Omron Sysmac Studio project SF_PLC ver.2 (Sysmac Studio 1.53.0.9, StandardProject)

# Controller new_controller_0: NX102-1020 version 1.33
Units and slaves: 노드1 : NX-ECC203 (E001); 유니트 1 : NX-ID6142-6 (N1); 유니트 2 : NX-OD6121-6 (N2); 유니트 1 : NX-PF0730 (N3); 유니트 2 : NX-ILM400 (N4); 유니트 4 : NX-SID800 (N6); 유니트 5 : NX-SOD400 (N7)
Task PrimaryTask (priority 4, period or condition 2000): Program0

TYPE Robot_IO : STRUCT
    IO : IO16;
END_STRUCT END_TYPE
TYPE IO16 : UNION
    w : WORD;
    b : ARRAY[1..32] OF BOOL;
END_UNION END_TYPE

VAR_GLOBAL
    Robot_In : ARRAY[0..237] OF WORD;  (* 로봇 > PLC; network input *)
    Robot_Out : ARRAY[0..105] OF WORD;  (* PLC > 로봇; network output *)
    vision_trig : BOOL;  (* 비전 촬영 신호; at ECAT://node#4/Line0 Trigger *)
    vis_data : DINT;  (* 비전 데이터; at ECAT://node#4/Line0 DINT Result Data 0 *)
    r_pause : BOOL;  (* 태스크 일시정지; at ECAT://node#[1,2]/Output Bit 32 bits/Output Bit 04 *)
    syl_f : BOOL;  (* 배출 실린더 전진; at ECAT://node#[1,2]/Output Bit 32 bits/Output Bit 05 *)
    syl_r : BOOL;  (* 배출 실린더 후진; at ECAT://node#[1,2]/Output Bit 32 bits/Output Bit 06 *)
    r_resume : BOOL;  (* 태스크 재개; at ECAT://node#[1,2]/Output Bit 32 bits/Output Bit 13 *)
    tower_R : BOOL;  (* 타워램프 - red; at ECAT://node#[1,2]/Output Bit 32 bits/Output Bit 20 *)
    tower_Y : BOOL;  (* 타워램프 - yellow; at ECAT://node#[1,2]/Output Bit 32 bits/Output Bit 21 *)
    tower_G : BOOL;  (* 타워램프 - green; at ECAT://node#[1,2]/Output Bit 32 bits/Output Bit 22 *)
    r_start : BOOL;  (* 태스크 실행; at ECAT://node#[1,2]/Output Bit 32 bits/Output Bit 23 *)
    r_stop : BOOL;  (* 태스크 정지; at ECAT://node#[1,2]/Output Bit 32 bits/Output Bit 24 *)
    vision_ss : BOOL;  (* 비전 감지 센서; at ECAT://node#[1,1]/Input Bit 32 bits/Input Bit 19 *)
    mag_ss : BOOL;  (* 매거진 센서; at ECAT://node#[1,1]/Input Bit 32 bits/Input Bit 23 *)
    stop_ss : BOOL;  (* 스토퍼 센서; at ECAT://node#[1,1]/Input Bit 32 bits/Input Bit 24 *)
    rsol_ss : BOOL;  (* 실린더 후진 센서; at ECAT://node#[1,1]/Input Bit 32 bits/Input Bit 25 *)
    fsol_ss : BOOL;  (* 실린더 전진 센서; at ECAT://node#[1,1]/Input Bit 32 bits/Input Bit 26 *)
    m_run : WORD;  (* 모터 구동; at ECAT://node#2/Command *)
    m_vel : UINT := 5000;  (* 모터 속도; at ECAT://node#2/Frequency reference *)
    m_status : WORD;  (* 모터 상태값; at ECAT://node#2/Status *)
    robot_recv : Robot_IO;  (* 로봇 I/O > PLC *)
    robot_send : Robot_IO;  (* PLC > 로봇 I/O *)
    robot_DI : Robot_IO;  (* 로봇 디지털 입력 *)
    manu_pb : BOOL;  (* 수동 운전 PB *)
    auto_pb : BOOL;  (* 자동 운전 PB *)
    f_sol_pb : BOOL;  (* 실린더 전진 PB *)
    r_sol_pb : BOOL;  (* 실린더 후진 PB *)
    conv_run : BOOL;  (* 모터 구동 PB *)
    conv_stop : BOOL;  (* 모터 정지 PB *)
    clamp_pb : BOOL;  (* 그리퍼 on *)
    uncalamp_pb : BOOL;  (* 그리퍼 off *)
    single_pb : BOOL;  (* 단속 동작 PB *)
    multi_pb : BOOL;  (* 연속 동작 PB *)
    count_val : INT;  (* 생산 수량 *)
    total_val : INT;  (* 적재부 *)
    save_val : INT;  (* 불량품 *)
    stop_pb : BOOL;  (* 정지 PB *)
    pause_pb : BOOL;  (* 일시정지 PB *)
    ems_pb : BOOL;  (* 비상 PB *)
    reset_pb : BOOL;  (* 리셋 PB *)
    places : ARRAY[1..6] OF BOOL;  (* 적재 상태 *)
    r_IO : ARRAY[1..7] OF WORD := [16#01, 16#02, 16#04, 16#08, 16#10, 16#20, 16#40];
    inductive_ss : BOOL;  (* 유도형 센서; at ECAT://node#[1,1]/Input Bit 32 bits/Input Bit 21 *)
    capacity_ss : BOOL;  (* 용량형 센서; at ECAT://node#[1,1]/Input Bit 32 bits/Input Bit 22 *)
    auto_busy : BOOL;
    manu_busy : BOOL;
    metal_cnt : INT;
    unmetal_cnt : INT;
END_VAR

(* Program Program0: safety or other program stored in binary form, left out *)

PROGRAM Program0
VAR
    task_on : BOOL;  (* 태스크 실행 신호 *)
    task_stop : BOOL;  (* 태스크 정지 신호 *)
    syl_f_manu : BOOL;  (* 수동 실린더 전진 *)
    syl_r_manu : BOOL;  (* 수동 실린더 후진 *)
    ready : BOOL;
    r_home : BOOL;  (* 로봇 홈 위치 *)
    single_busy : BOOL;
    multi_busy : BOOL;
    mps_start : BOOL;
    m_step : INT;
    stop_act : BOOL;
    pause_act : BOOL;
    resume_act : BOOL;
    resume_T : TON;
    resume_T1 : TON;
    pause_T1 : TON;
    pause_T2 : TON;
    red_a : BOOL;
    red_b : BOOL;
    ems_act : BOOL;
    reset_act : BOOL;
    reset_T : TON;
    reset_all : BOOL;
    syl_r_auto : BOOL;  (* 실린더 상태 리셋 *)
    syl_f_mps : BOOL;  (* 자동 실린더 전진 *)
    syl_r_mps : BOOL;  (* 자동 실린더 후진 *)
    vision_T : TON;
    vis_no : DINT;
    robot_start : BOOL;
    mps_busy : BOOL;
    r_step : INT;
    robot_busy : BOOL;
    r_status : WORD;
    r_done : BOOL;  (* 로봇 done *)
    robot_done : BOOL;
    counter : CTU;
    cnt_reset : BOOL;
    retry : BOOL;
    grip_close : BOOL;  (* 그리퍼 on *)
    grip_open : BOOL;  (* 그리퍼 off *)
    tast_T : TON;
    metal_ss : BOOL;
END_VAR
VAR_EXTERNAL
    robot_recv : Robot_IO;
    robot_send : Robot_IO;
    Robot_Out : ARRAY[0..105] OF WORD;
    Robot_In : ARRAY[0..237] OF WORD;
    robot_DI : Robot_IO;
    manu_pb : BOOL;
    auto_pb : BOOL;
    r_start : BOOL;
    r_stop : BOOL;
    f_sol_pb : BOOL;
    m_run : WORD;
    r_sol_pb : BOOL;
    conv_run : BOOL;
    conv_stop : BOOL;
    clamp_pb : BOOL;
    uncalamp_pb : BOOL;
    mag_ss : BOOL;
    rsol_ss : BOOL;
    single_pb : BOOL;
    multi_pb : BOOL;
    count_val : INT;
    vis_data : DINT;
    stop_pb : BOOL;
    pause_pb : BOOL;
    r_pause : BOOL;
    r_resume : BOOL;
    tower_R : BOOL;
    ems_pb : BOOL;
    reset_pb : BOOL;
    syl_r : BOOL;
    syl_f : BOOL;
    places : ARRAY[1..6] OF BOOL;
    m_status : WORD;
    total_val : INT;
    save_val : INT;
    fsol_ss : BOOL;
    vision_ss : BOOL;
    stop_ss : BOOL;
    vision_trig : BOOL;
    r_IO : ARRAY[1..7] OF WORD;
    tower_Y : BOOL;
    tower_G : BOOL;
    auto_busy : BOOL;
    manu_busy : BOOL;
    capacity_ss : BOOL;
    inductive_ss : BOOL;
    metal_cnt : INT;
    unmetal_cnt : INT;
END_VAR
VAR
    _e1 : F_TRIG;
    _e2 : R_TRIG;
    _e3 : R_TRIG;
    _p4 : BOOL;
    _e5 : R_TRIG;
    _e6 : R_TRIG;
    _e7 : R_TRIG;
    _p8 : BOOL;
    _e9 : F_TRIG;
    _e10 : R_TRIG;
    _e11 : R_TRIG;
    _e12 : F_TRIG;
END_VAR

(* Section comm: ladder, written here as Structured Text *)

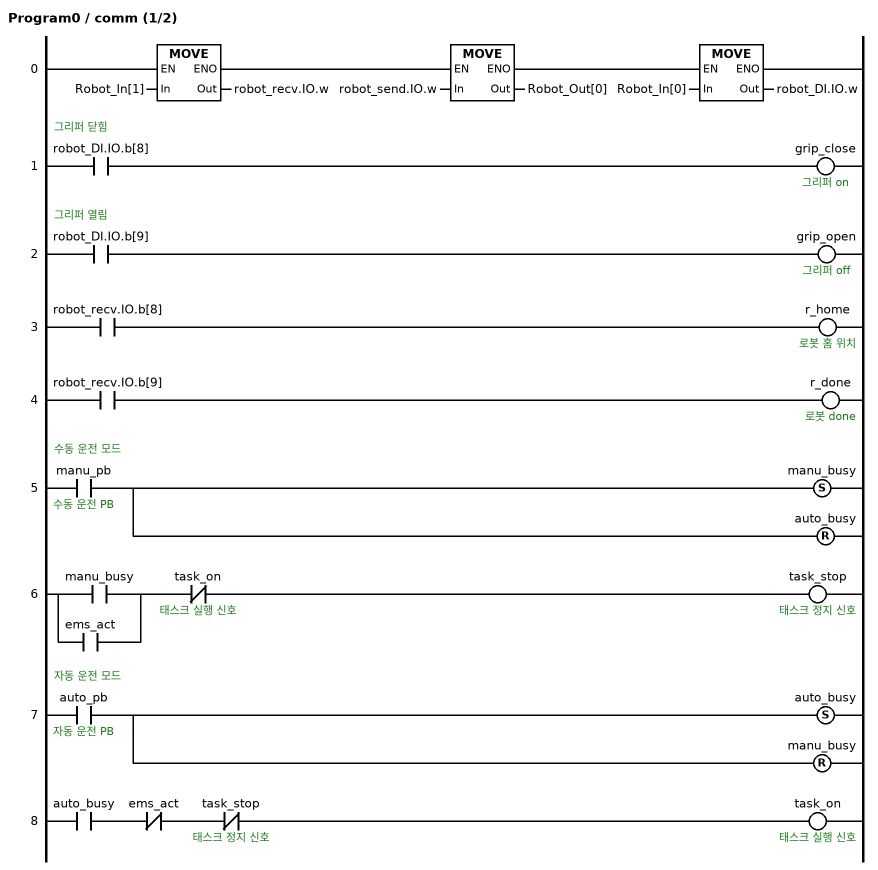
(* Rung 0 *)
robot_recv.IO.w := Robot_In[1];
Robot_Out[0] := robot_send.IO.w;
robot_DI.IO.w := Robot_In[0];
(* Rung 1: 그리퍼 닫힘 *)
grip_close := robot_DI.IO.b[8];
(* Rung 2: 그리퍼 열림 *)
grip_open := robot_DI.IO.b[9];
(* Rung 3 *)
r_home := robot_recv.IO.b[8];
(* Rung 4 *)
r_done := robot_recv.IO.b[9];
(* Rung 5: 수동 운전 모드 *)
IF manu_pb THEN
    manu_busy := TRUE;
    auto_busy := FALSE;
END_IF;
(* Rung 6 *)
task_stop := (manu_busy OR ems_act) AND NOT task_on;
(* Rung 7: 자동 운전 모드 *)
IF auto_pb THEN
    auto_busy := TRUE;
    manu_busy := FALSE;
END_IF;
(* Rung 8 *)
task_on := auto_busy AND NOT ems_act AND NOT task_stop;

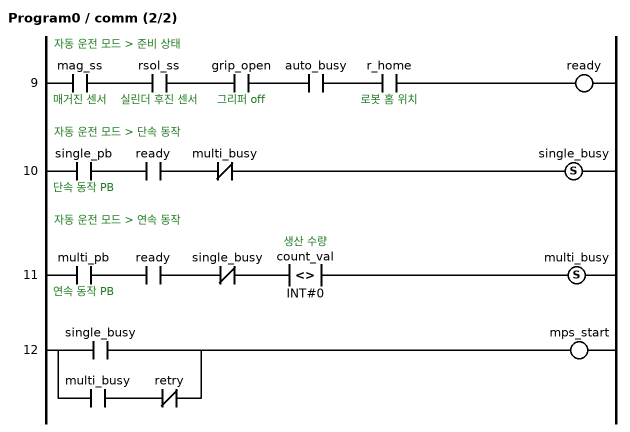
(* Rung 9: 자동 운전 모드 > 준비 상태 *)
ready := mag_ss AND rsol_ss AND grip_open AND auto_busy AND r_home;
(* Rung 10: 자동 운전 모드 > 단속 동작 *)
IF single_pb AND ready AND NOT multi_busy THEN single_busy := TRUE; END_IF;
(* Rung 11: 자동 운전 모드 > 연속 동작 *)
IF multi_pb AND ready AND NOT single_busy AND (count_val <> INT#0) THEN multi_busy := TRUE; END_IF;
(* Rung 12 *)
mps_start := single_busy OR (multi_busy AND NOT retry);

(* Section manual: ladder, written here as Structured Text *)

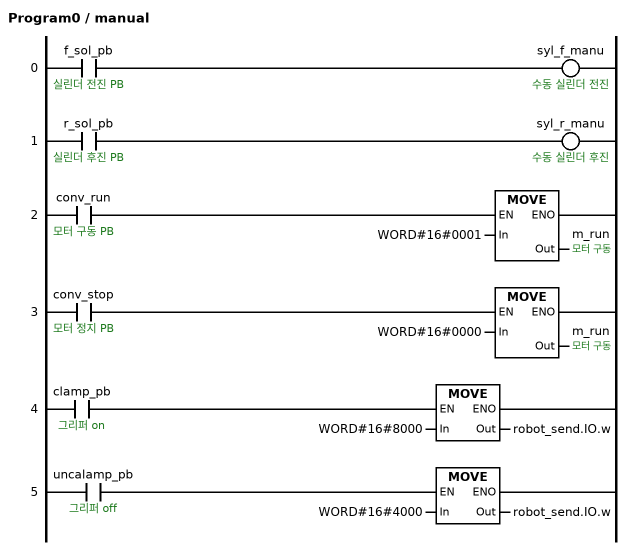
(* Rung 0 *)
syl_f_manu := f_sol_pb;
(* Rung 1 *)
syl_r_manu := r_sol_pb;
(* Rung 2 *)
IF conv_run THEN m_run := WORD#16#0001; END_IF;
(* Rung 3 *)
IF conv_stop THEN m_run := WORD#16#0000; END_IF;
(* Rung 4 *)
IF clamp_pb THEN robot_send.IO.w := WORD#16#8000; END_IF;
(* Rung 5 *)
IF uncalamp_pb THEN robot_send.IO.w := WORD#16#4000; END_IF;

(* Section auto: ladder, written here as Structured Text *)

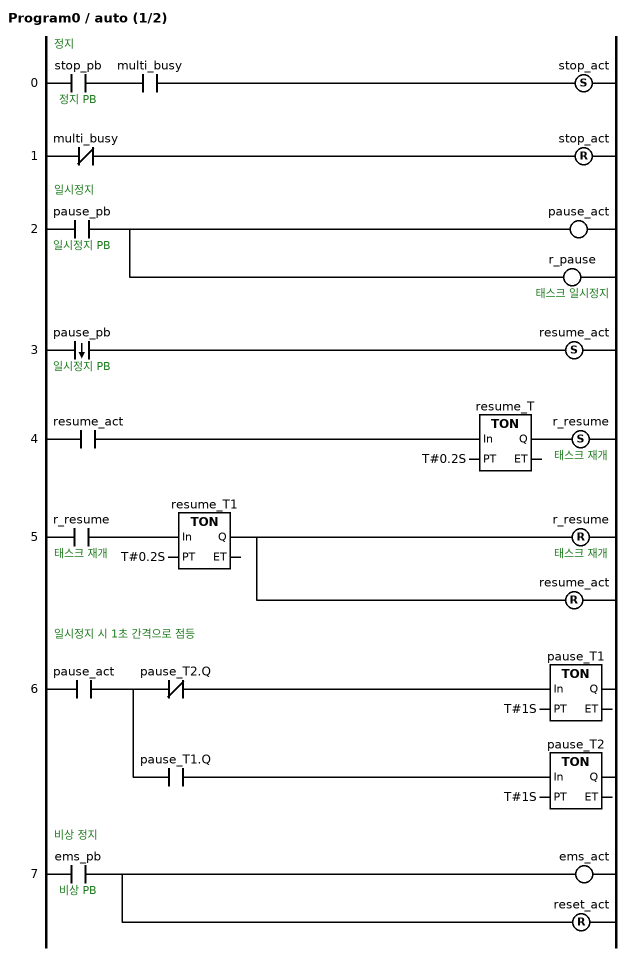
(* Rung 0: 정지 *)
IF stop_pb AND multi_busy THEN stop_act := TRUE; END_IF;
(* Rung 1 *)
IF NOT multi_busy THEN stop_act := FALSE; END_IF;
(* Rung 2: 일시정지 *)
pause_act := pause_pb;
r_pause := pause_pb;
(* Rung 3 *)
_e1(CLK := pause_pb);
IF _e1.Q THEN resume_act := TRUE; END_IF;
(* Rung 4 *)
resume_T(In := resume_act, PT := T#0.2S);
IF resume_T.Q THEN r_resume := TRUE; END_IF;
(* Rung 5 *)
resume_T1(In := r_resume, PT := T#0.2S);
IF resume_T1.Q THEN
    r_resume := FALSE;
    resume_act := FALSE;
END_IF;
(* Rung 6: 일시정지 시 1초 간격으로 점등 *)
pause_T1(In := pause_act AND NOT pause_T2.Q, PT := T#1S);
pause_T2(In := pause_act AND pause_T1.Q, PT := T#1S);
(* Rung 7: 비상 정지 *)
ems_act := ems_pb;
IF ems_pb THEN reset_act := FALSE; END_IF;

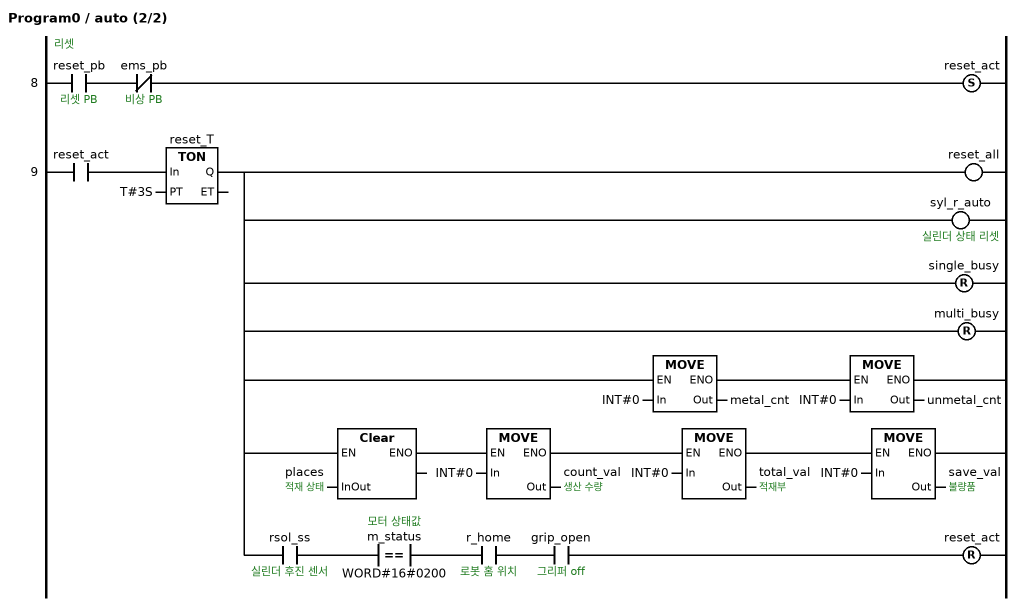
(* Rung 8: 리셋 *)
IF reset_pb AND NOT ems_pb THEN reset_act := TRUE; END_IF;
(* Rung 9 *)
reset_T(In := reset_act, PT := T#3S);
reset_all := reset_T.Q;
syl_r_auto := reset_T.Q;
IF reset_T.Q THEN
    single_busy := FALSE;
    multi_busy := FALSE;
    metal_cnt := INT#0;
    unmetal_cnt := INT#0;
    Clear(InOut := places);
    count_val := INT#0;
    total_val := INT#0;
    save_val := INT#0;
END_IF;
IF reset_T.Q AND rsol_ss AND (m_status = WORD#16#0200) AND r_home AND grip_open THEN
    reset_act := FALSE;
END_IF;

(* Section mps: ladder, written here as Structured Text *)

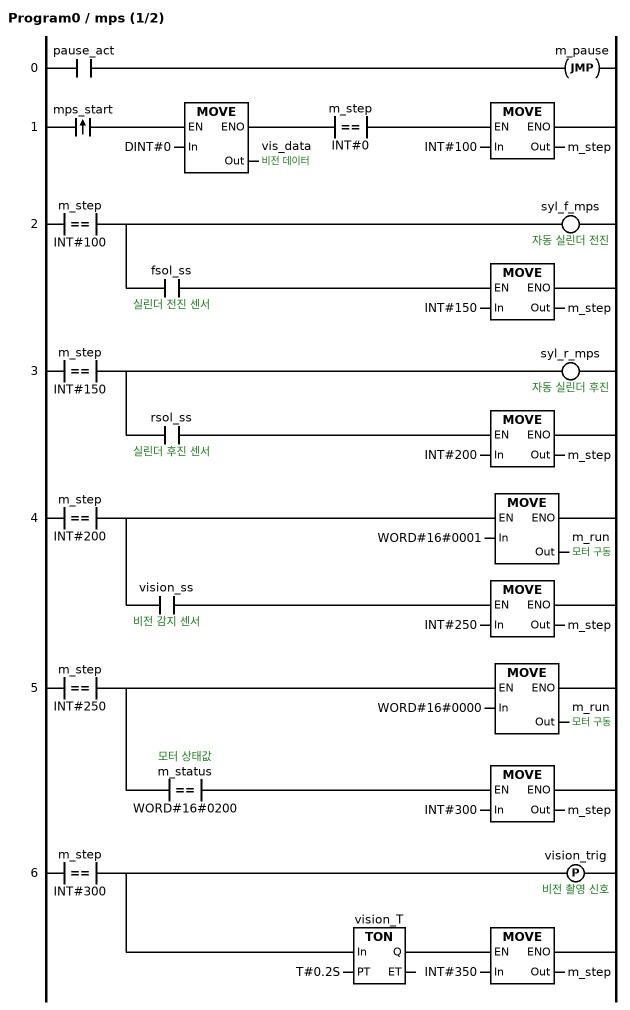
(* Rung 0 *)
IF pause_act THEN JMP m_pause; END_IF;
(* Rung 1 *)
_e2(CLK := mps_start);
IF _e2.Q THEN vis_data := DINT#0; END_IF;
IF _e2.Q AND (m_step = INT#0) THEN m_step := INT#100; END_IF;
(* Rung 2 *)
syl_f_mps := m_step = INT#100;
IF (m_step = INT#100) AND fsol_ss THEN m_step := INT#150; END_IF;
(* Rung 3 *)
syl_r_mps := m_step = INT#150;
IF (m_step = INT#150) AND rsol_ss THEN m_step := INT#200; END_IF;
(* Rung 4 *)
IF m_step = INT#200 THEN m_run := WORD#16#0001; END_IF;
IF (m_step = INT#200) AND vision_ss THEN m_step := INT#250; END_IF;
(* Rung 5 *)
IF m_step = INT#250 THEN m_run := WORD#16#0000; END_IF;
IF (m_step = INT#250) AND (m_status = WORD#16#0200) THEN m_step := INT#300; END_IF;
(* Rung 6 *)
_e3(CLK := m_step = INT#300);
vision_trig := _e3.Q;
vision_T(In := m_step = INT#300, PT := T#0.2S);
IF vision_T.Q THEN m_step := INT#350; END_IF;

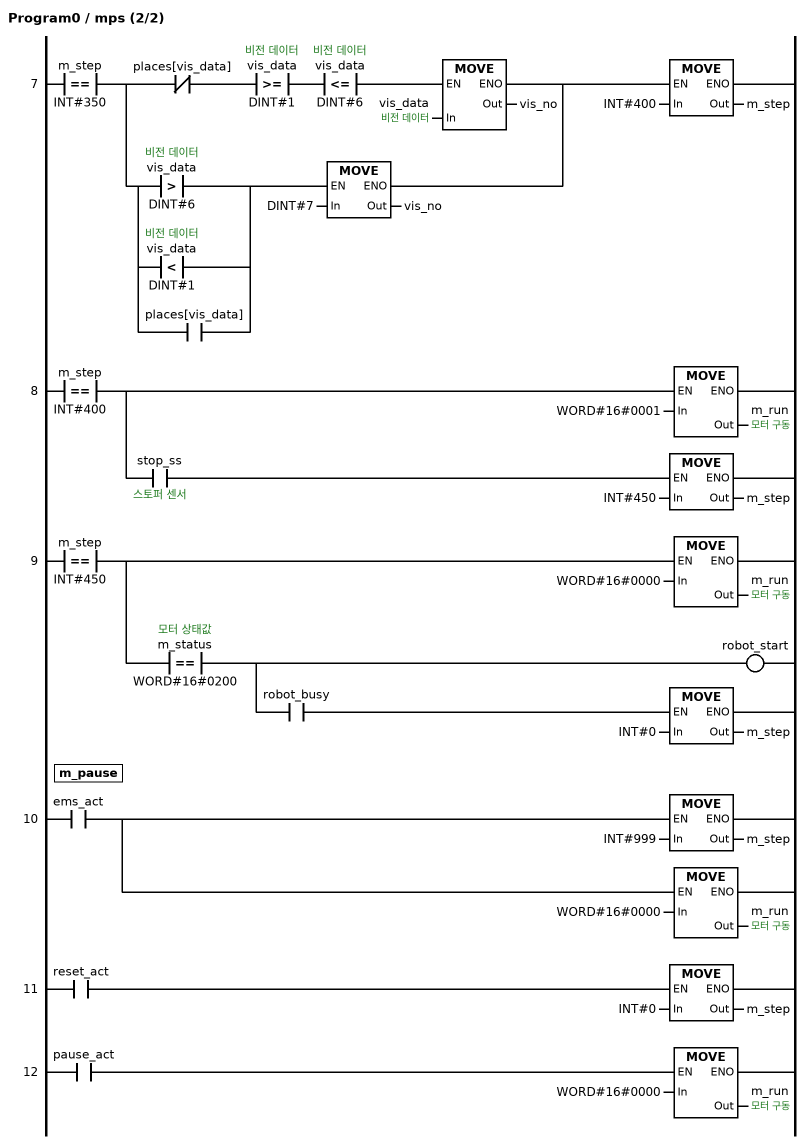
(* Rung 7 *)
IF (m_step = INT#350) AND NOT places[vis_data] AND (vis_data >= DINT#1) AND (vis_data <= DINT#6) THEN
    vis_no := vis_data;
END_IF;
IF (m_step = INT#350) AND ((vis_data > DINT#6) OR (vis_data < DINT#1) OR places[vis_data]) THEN
    vis_no := DINT#7;
END_IF;
IF (m_step = INT#350) AND ((NOT places[vis_data] AND (vis_data >= DINT#1) AND (vis_data <= DINT#6)) OR (vis_data > DINT#6) OR (vis_data < DINT#1) OR places[vis_data]) THEN
    m_step := INT#400;
END_IF;
(* Rung 8 *)
IF m_step = INT#400 THEN m_run := WORD#16#0001; END_IF;
IF (m_step = INT#400) AND stop_ss THEN m_step := INT#450; END_IF;
(* Rung 9 *)
IF m_step = INT#450 THEN m_run := WORD#16#0000; END_IF;
robot_start := (m_step = INT#450) AND (m_status = WORD#16#0200);
IF (m_step = INT#450) AND (m_status = WORD#16#0200) AND robot_busy THEN m_step := INT#0; END_IF;
(* Rung 10 *)
m_pause:
IF ems_act THEN
    m_step := INT#999;
    m_run := WORD#16#0000;
END_IF;
(* Rung 11 *)
IF reset_act THEN m_step := INT#0; END_IF;
(* Rung 12 *)
IF pause_act THEN m_run := WORD#16#0000; END_IF;

(* Section robot: ladder, written here as Structured Text *)

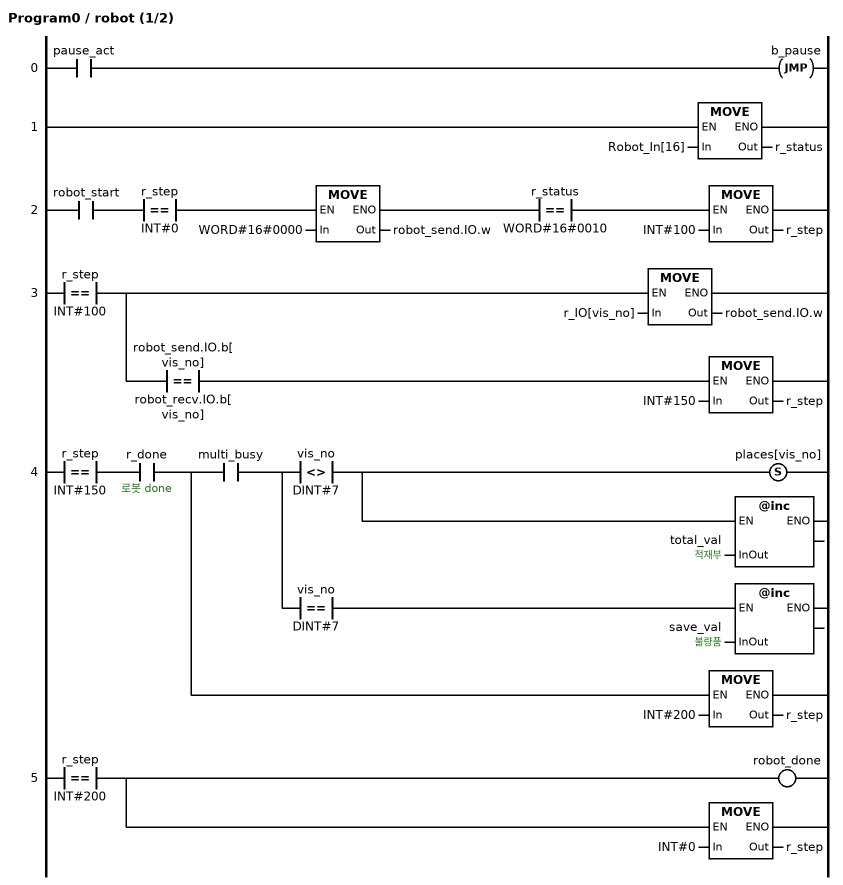
(* Rung 0 *)
IF pause_act THEN JMP b_pause; END_IF;
(* Rung 1 *)
r_status := Robot_In[16];
(* Rung 2 *)
IF robot_start AND (r_step = INT#0) THEN robot_send.IO.w := WORD#16#0000; END_IF;
IF robot_start AND (r_step = INT#0) AND (r_status = WORD#16#0010) THEN r_step := INT#100; END_IF;
(* Rung 3 *)
IF r_step = INT#100 THEN robot_send.IO.w := r_IO[vis_no]; END_IF;
IF (r_step = INT#100) AND (robot_send.IO.b[vis_no] = robot_recv.IO.b[vis_no]) THEN
    r_step := INT#150;
END_IF;
(* Rung 4 *)
_p4 := (r_step = INT#150) AND r_done AND multi_busy AND (vis_no <> DINT#7);
IF _p4 THEN places[vis_no] := TRUE; END_IF;
_e5(CLK := _p4);
IF _e5.Q THEN inc(InOut := total_val); END_IF;
_e6(CLK := (r_step = INT#150) AND r_done AND multi_busy AND (vis_no = DINT#7));
IF _e6.Q THEN inc(InOut := save_val); END_IF;
IF (r_step = INT#150) AND r_done THEN r_step := INT#200; END_IF;
(* Rung 5 *)
robot_done := r_step = INT#200;
IF r_step = INT#200 THEN r_step := INT#0; END_IF;

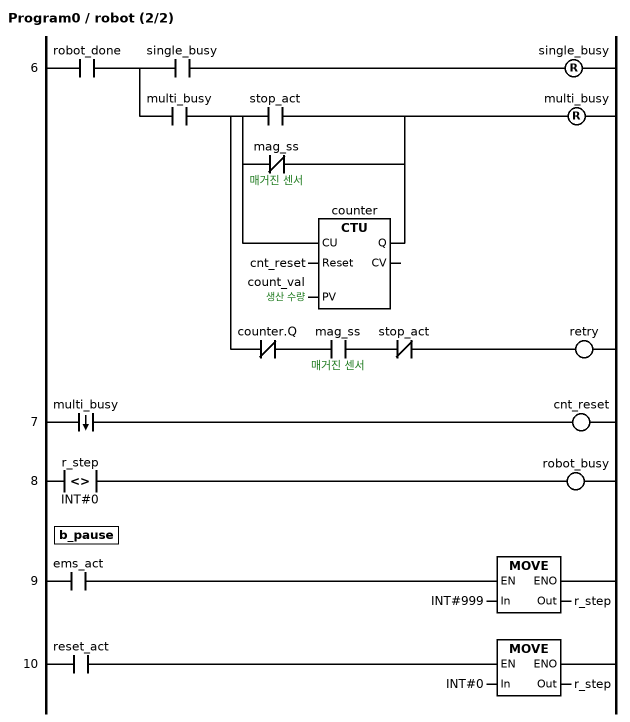
(* Rung 6 *)
IF robot_done AND single_busy THEN single_busy := FALSE; END_IF;
_e7(CLK := robot_done AND multi_busy);
counter(CU := _e7.Q, Reset := cnt_reset, PV := count_val);
_p8 := robot_done AND multi_busy;
IF (robot_done AND multi_busy AND (stop_act OR NOT mag_ss)) OR counter.Q THEN multi_busy := FALSE; END_IF;
retry := _p8 AND NOT counter.Q AND mag_ss AND NOT stop_act;
(* Rung 7 *)
_e9(CLK := multi_busy);
cnt_reset := _e9.Q;
(* Rung 8 *)
robot_busy := r_step <> INT#0;
(* Rung 9 *)
b_pause:
IF ems_act THEN r_step := INT#999; END_IF;
(* Rung 10 *)
IF reset_act THEN r_step := INT#0; END_IF;

(* Section output: ladder, written here as Structured Text *)

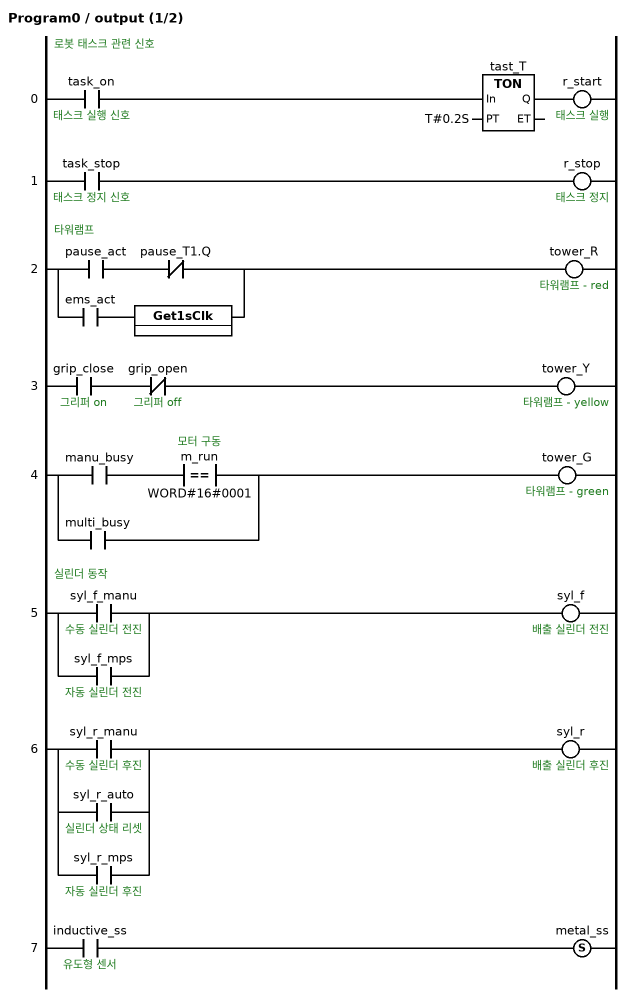
(* Rung 0: 로봇 태스크 관련 신호 *)
tast_T(In := task_on, PT := T#0.2S);
r_start := tast_T.Q;
(* Rung 1 *)
r_stop := task_stop;
(* Rung 2: 타워램프 *)
tower_R := (pause_act AND NOT pause_T1.Q) OR (ems_act AND Get1sClk());
(* Rung 3 *)
tower_Y := grip_close AND NOT grip_open;
(* Rung 4 *)
tower_G := (manu_busy AND (m_run = WORD#16#0001)) OR multi_busy;
(* Rung 5: 실린더 동작 *)
syl_f := syl_f_manu OR syl_f_mps;
(* Rung 6 *)
syl_r := syl_r_manu OR syl_r_auto OR syl_r_mps;
(* Rung 7 *)
IF inductive_ss THEN metal_ss := TRUE; END_IF;

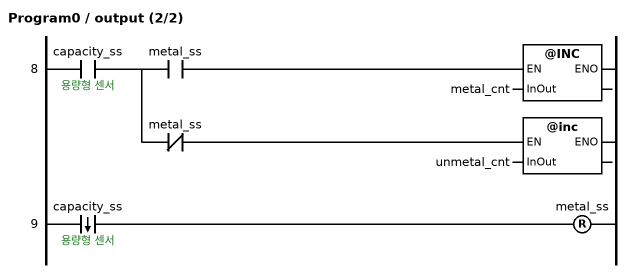
(* Rung 8 *)
_e10(CLK := capacity_ss AND metal_ss);
IF _e10.Q THEN INC(InOut := metal_cnt); END_IF;
_e11(CLK := capacity_ss AND NOT metal_ss);
IF _e11.Q THEN inc(InOut := unmetal_cnt); END_IF;
(* Rung 9 *)
_e12(CLK := capacity_ss);
IF _e12.Q THEN metal_ss := FALSE; END_IF;
END_PROGRAM

# Device HMI_NA5_0 (NA): not converted